// TIA Portal V17 export
// export: Created 2026-11-10T15:00:48.6641979Z, ExportSetting WithDefaults, DisplayName Totally Integrated Automation Portal, DisplayVersion V17, DisplayName TIA Portal Openness, DisplayVersion V17, DisplayName TIA Portal Version Control Interface, DisplayVersion V17, DisplayName STEP 7 Professional, DisplayVersion V17, DisplayName STEP 7 Safety, DisplayVersion V17, DisplayName WinCC Advanced, DisplayVersion V17
GraphicList "Level120"  ListRange=Decimal, Mode=Simple
  GraphicListEntry   EntryType=Range, To=11, Picture=Tank_0
  GraphicListEntry   EntryType=Range, From=12, To=23, Picture=Tank_1
  GraphicListEntry   EntryType=Range, From=24, To=35, Picture=Tank_2
  GraphicListEntry   EntryType=Range, From=36, To=47, Picture=Tank_3
  GraphicListEntry   EntryType=Range, From=48, To=59, Picture=Tank_4
  GraphicListEntry   EntryType=Range, From=60, To=71, Picture=Tank_5
  GraphicListEntry   EntryType=Range, From=72, To=83, Picture=Tank_6
  GraphicListEntry   EntryType=Range, From=84, To=95, Picture=Tank_7
  GraphicListEntry   EntryType=Range, From=96, To=107, Picture=Tank_8
  GraphicListEntry   EntryType=Range, From=108, To=119, Picture=Tank_9
  GraphicListEntry   EntryType=Range, From=120, To=120, Picture=Tank_10
